Staubli VAL3: resizeMark.pgx

public program resizeMark(string x_sKey)
  local num l_nSize
  local num l_i
begin
  call getPointSize(x_sKey,l_nSize)
  //resize(savedata:nMarkIndex,1,l_nSize)
  for l_i = 0 to l_nSize-1
    trajTemp:tTrajItem[x_sKey].pPointItem[l_i].bMarked=false
  endFor
end
